(* CODESYS project P_ClassName.xml

Project tree, tasks and I/O mapping:
*)

// P_ClassName
PROPERTY P_ClassName : STRING
END_PROPERTY
